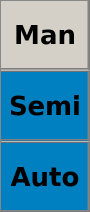
VISUALIZATION Mode_Select_1  // 90x212
VAR_IN_OUT
	stMode: ST_Mode;
END_VAR
    Button (0,0 90x70), "Man", colour toggle: stModeMain.iActMode=eManualMode, input disabled if: NOT GVL.MainMachine.bReadyToManualModeSelect
        OnMouseDown: execute {
            stModeMain.bSetManual:=TRUE;
            stMode.bSetSemi:=FALSE;
            stMode.bSetAuto:=FALSE;
        }
    Button (0,71 90x70), "Semi", colour toggle: stModeMain.iActMode=eSemiAutoMode, input disabled if: stModeMain.iActMode<>E_WorkingMode.eManualMode
        OnMouseDown: execute {
            stModeMain.bSetManual:=FALSE;
            stMode.bSetSemi:=TRUE;
            stMode.bSetAuto:=FALSE;
        }
    Button (0,142 90x70), "Auto", colour toggle: stModeMain.iActMode=eAutoMode, input disabled if: stModeMain.iActMode<>E_WorkingMode.eManualMode
        OnMouseDown: execute {
            stModeMain.bSetManual:=FALSE;
            stMode.bSetSemi:=FALSE;
            stMode.bSetAuto:=TRUE;
        }
END_VISUALIZATION

(* stored: Version 1.1.0.1, ProductVersion 3.1.4024.13
   Visu Mode_Select_1: Id {73246c8e-1504-4fe9-b4c8-76699e009a9f} *)
